TYPE "ST_SequenceCursor"
VERSION : 0.1
   STRUCT
      RowIdx : Int;
      Elapsed : Time;
      TimedOut : Bool;
   END_STRUCT;

END_TYPE

